Fanuc KAREL source: compact_preamble.KL

PROGRAM KT00893
%NOLOCKGROUP
VAR
P1 : POSITION;P2 : POSITION;OUT:BOOLEAN
BEGIN
OUT=IN_RANGE(P1)
END KT00893
